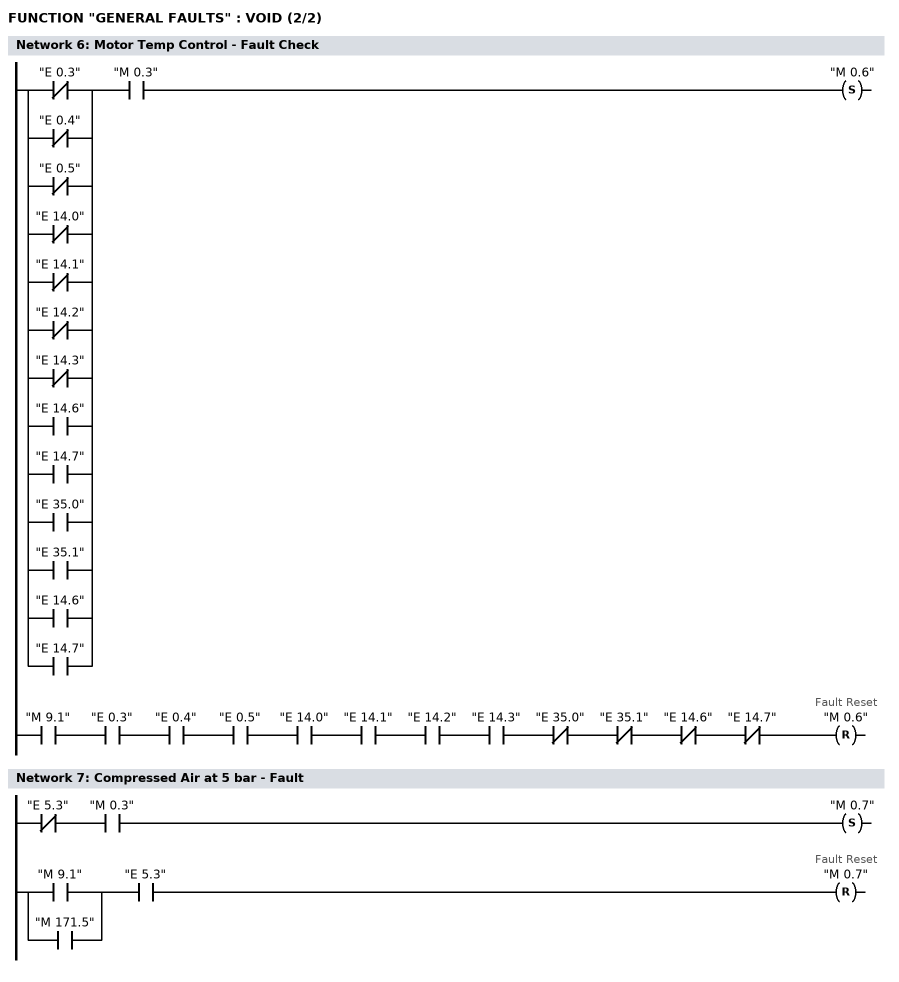

      A(    ;
      ON    "E 0.3";
      ON    "E 0.4";
      ON    "E 0.5";
      ON    "E 14.0";
      ON    "E 14.1";
      ON    "E 14.2";
      ON    "E 14.3";
      O     "E 14.6";
      O     "E 14.7";
      O     "E 35.0";
      O     "E 35.1";
      O     "E 14.6";
      O     "E 14.7";
      )     ;
      A     "M 0.3";
      S     "M 0.6";
//;
      A     "M 9.1";
      A     "E 0.3";
      A     "E 0.4";
      A     "E 0.5";
      A     "E 14.0";
      A     "E 14.1";
      A     "E 14.2";
      A     "E 14.3";
      AN    "E 35.0";
      AN    "E 35.1";
      AN    "E 14.6";
      AN    "E 14.7";
      R     "M 0.6"; // Fault Reset
NETWORK
TITLE =Compressed Air at 5 bar - Fault

      AN    "E 5.3";
      A     "M 0.3";
      S     "M 0.7";
//;
      A(    ;
      O     "M 9.1";
      O     "M 171.5";
      )     ;
      A     "E 5.3";
      R     "M 0.7"; // Fault Reset
NETWORK
TITLE =Faults Register 1 - E-Stops & Safety Doors

      A(    ;
      L     "MB 1";
      L     0;
      <>I   ;
      )     ;
      =     #FAULT_REGISTER_1;
//;
      A     #FAULT_REGISTER_1;
      O     #CHECK_PULSE;
      O     "M 17.1";
      O     "M 9.1";
      JNB   FR01;
NETWORK
TITLE =E-Stop  Desk  X120
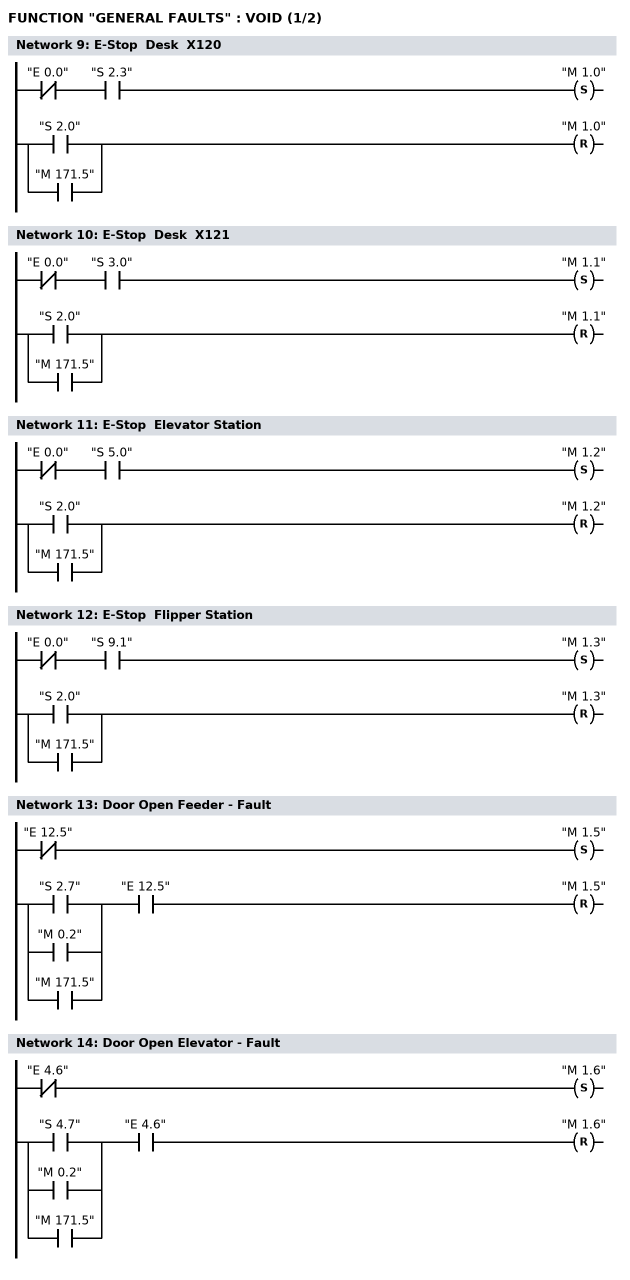

      AN    "E 0.0";
      A     "S 2.3";
      S     "M 1.0";
//;
      A(    ;
      O     "S 2.0";
      O     "M 171.5";
      )     ;
      R     "M 1.0";
NETWORK
TITLE =E-Stop  Desk  X121

      AN    "E 0.0";
      A     "S 3.0";
      S     "M 1.1";
//;
      A(    ;
      O     "S 2.0";
      O     "M 171.5";
      )     ;
      R     "M 1.1";
NETWORK
TITLE =E-Stop  Elevator Station

      AN    "E 0.0";
      A     "S 5.0";
      S     "M 1.2";
//;
      A(    ;
      O     "S 2.0";
      O     "M 171.5";
      )     ;
      R     "M 1.2";
NETWORK
TITLE =E-Stop  Flipper Station

      AN    "E 0.0";
      A     "S 9.1";
      S     "M 1.3";
//;
      A(    ;
      O     "S 2.0";
      O     "M 171.5";
      )     ;
      R     "M 1.3";
NETWORK
TITLE =Door Open Feeder - Fault

      AN    "E 12.5";
      S     "M 1.5";
//;
      A(    ;
      O     "S 2.7";
      O     "M 0.2";
      O     "M 171.5";
      )     ;
      A     "E 12.5";
      R     "M 1.5";
NETWORK
TITLE =Door Open Elevator - Fault

      AN    "E 4.6";
      S     "M 1.6";
//;
      A(    ;
      O     "S 4.7";
      O     "M 0.2";
      O     "M 171.5";
      )     ;
      A     "E 4.6";
      R     "M 1.6";
NETWORK
TITLE =Door Open Flipper - Fault
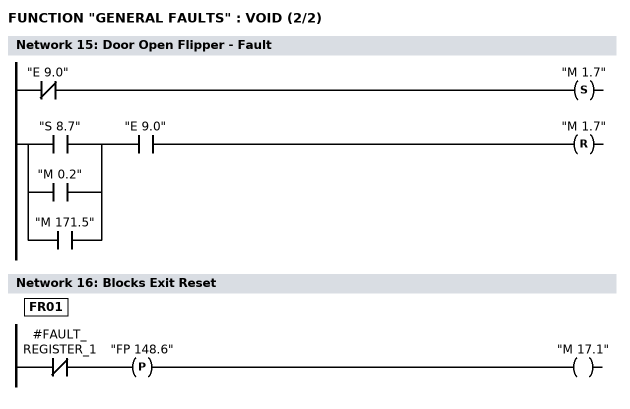

      AN    "E 9.0";
      S     "M 1.7";
//;
      A(    ;
      O     "S 8.7";
      O     "M 0.2";
      O     "M 171.5";
      )     ;
      A     "E 9.0";
      R     "M 1.7";
NETWORK
TITLE =Blocks Exit Reset

FR01: NOP   0;

      AN    #FAULT_REGISTER_1;
      FP    "FP 148.6";
      =     "M 17.1";
NETWORK
TITLE =Faults Register 2 - Conveyor 0 to Conveyor 3

      A(    ;
      L     "MB 2";
      L     0;
      <>I   ;
      )     ;
      =     #FAULT_REGISTER_2;
      =     "HMI_DB".SCREEN_CALL_1;
//;
      A     #FAULT_REGISTER_2;
      O     #CHECK_PULSE;
      O     "M 17.2";
      O     "M 9.1";
      JNB   FR02;
NETWORK
TITLE =K62.0 / 1 Conveyor 0 - Fault
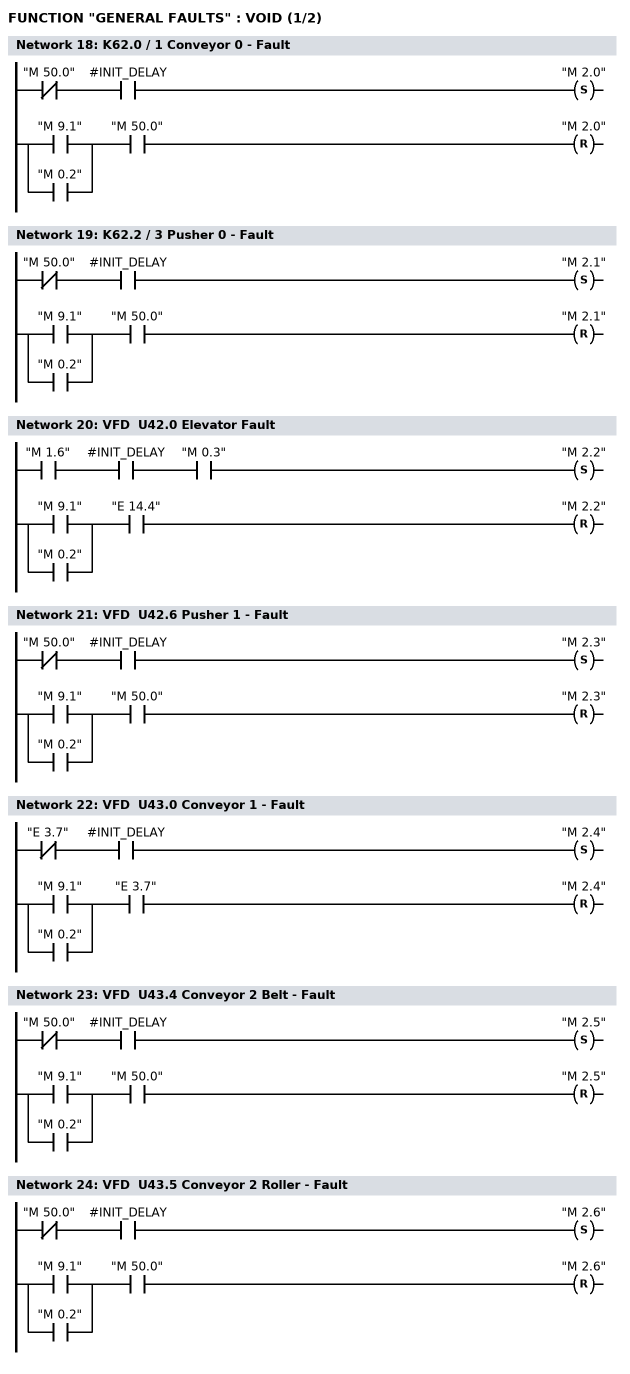

      AN    "M 50.0";
      A     #INIT_DELAY;
      S     "M 2.0";
//;
      A(    ;
      O     "M 9.1";
      O     "M 0.2";
      )     ;
      A     "M 50.0";
      R     "M 2.0";
NETWORK
TITLE =K62.2 / 3 Pusher 0 - Fault

      AN    "M 50.0";
      A     #INIT_DELAY;
      S     "M 2.1";
//;
      A(    ;
      O     "M 9.1";
      O     "M 0.2";
      )     ;
      A     "M 50.0";
      R     "M 2.1";
NETWORK
TITLE =VFD  U42.0 Elevator Fault

//   AN    #ELEVATOR_U42_0
      A     "M 1.6";
      A     #INIT_DELAY;
      A     "M 0.3";
      S     "M 2.2";
//;
      A(    ;
      O     "M 9.1";
      O     "M 0.2";
      )     ;
//      A     "E 3.6"
      A     "E 14.4";
      R     "M 2.2";
NETWORK
TITLE =VFD  U42.6 Pusher 1 - Fault

      AN    "M 50.0";
      A     #INIT_DELAY;
      S     "M 2.3";
//;
      A(    ;
      O     "M 9.1";
      O     "M 0.2";
      )     ;
      A     "M 50.0";
      R     "M 2.3";
NETWORK
TITLE =VFD  U43.0 Conveyor 1 - Fault

      AN    "E 3.7";
      A     #INIT_DELAY;
      S     "M 2.4";
//;
      A(    ;
      O     "M 9.1";
      O     "M 0.2";
      )     ;
      A     "E 3.7";
      R     "M 2.4";
NETWORK
TITLE =VFD  U43.4 Conveyor 2 Belt - Fault

      AN    "M 50.0";
      A     #INIT_DELAY;
      S     "M 2.5";
//;
      A(    ;
      O     "M 9.1";
      O     "M 0.2";
      )     ;
      A     "M 50.0";
      R     "M 2.5";
NETWORK
TITLE =VFD  U43.5 Conveyor 2 Roller - Fault

      AN    "M 50.0";
      A     #INIT_DELAY;
      S     "M 2.6";
//;
      A(    ;
      O     "M 9.1";
      O     "M 0.2";
      )     ;
      A     "M 50.0";
      R     "M 2.6";
NETWORK
TITLE =VFD  U44.0 Conveyor 3 Fault
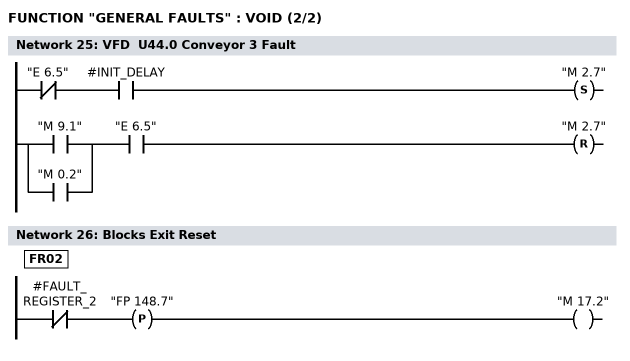

      AN    "E 6.5";
      A     #INIT_DELAY;
      S     "M 2.7";
//;
      A(    ;
      O     "M 9.1";
      O     "M 0.2";
      )     ;
      A     "E 6.5";
      R     "M 2.7";
NETWORK
TITLE =Blocks Exit Reset

FR02: NOP   0;

      AN    #FAULT_REGISTER_2;
      FP    "FP 148.7";
      =     "M 17.2";
NETWORK
TITLE =Faults Register 3 - Conveyor 4 to Conveyor 9

      A(    ;
      L     "MB 3";
      L     0;
      <>I   ;
      )     ;
      =     #FAULT_REGISTER_3;
      =     "HMI_DB".SCREEN_CALL_2;
//;
      A     #FAULT_REGISTER_3;
      O     #CHECK_PULSE;
      O     "M 17.3";
      O     "M 9.1";
      JNB   FR03;
NETWORK
TITLE =VFD  U44.3 Fault
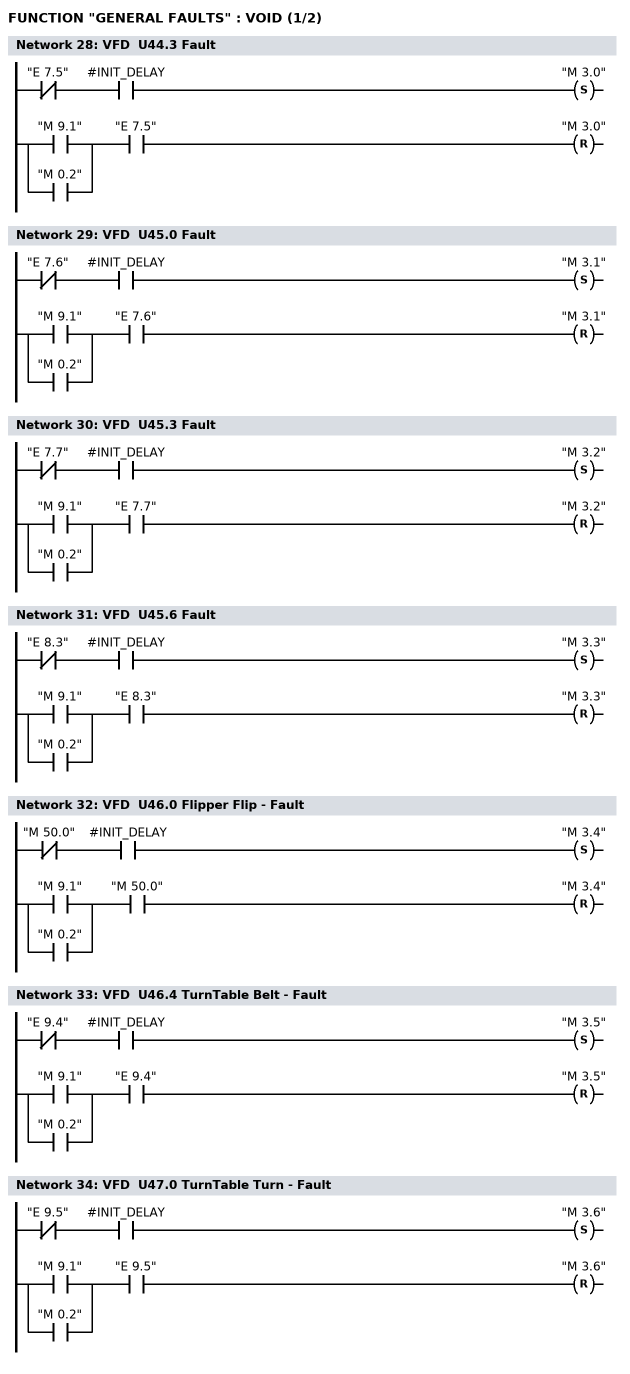

      AN    "E 7.5";
      A     #INIT_DELAY;
      S     "M 3.0";
//;
      A(    ;
      O     "M 9.1";
      O     "M 0.2";
      )     ;
      A     "E 7.5";
      R     "M 3.0";
NETWORK
TITLE =VFD  U45.0 Fault

      AN    "E 7.6";
      A     #INIT_DELAY;
      S     "M 3.1";
//;
      A(    ;
      O     "M 9.1";
      O     "M 0.2";
      )     ;
      A     "E 7.6";
      R     "M 3.1";
NETWORK
TITLE =VFD  U45.3 Fault

      AN    "E 7.7";
      A     #INIT_DELAY;
      S     "M 3.2";
//;
      A(    ;
      O     "M 9.1";
      O     "M 0.2";
      )     ;
      A     "E 7.7";
      R     "M 3.2";
NETWORK
TITLE =VFD  U45.6 Fault

      AN    "E 8.3";
      A     #INIT_DELAY;
      S     "M 3.3";
///;
      A(    ;
      O     "M 9.1";
      O     "M 0.2";
      )     ;
      A     "E 8.3";
      R     "M 3.3";
NETWORK
TITLE =VFD  U46.0 Flipper Flip - Fault

      AN    "M 50.0";
      A     #INIT_DELAY;
      S     "M 3.4";
//;
      A(    ;
      O     "M 9.1";
      O     "M 0.2";
      )     ;
      A     "M 50.0";
      R     "M 3.4";
NETWORK
TITLE =VFD  U46.4 TurnTable Belt - Fault

      AN    "E 9.4";
      A     #INIT_DELAY;
      S     "M 3.5";
//;
      A(    ;
      O     "M 9.1";
      O     "M 0.2";
      )     ;
      A     "E 9.4";
      R     "M 3.5";
NETWORK
TITLE =VFD  U47.0 TurnTable Turn - Fault

      AN    "E 9.5";
      A     #INIT_DELAY;
      S     "M 3.6";
//;
      A(    ;
      O     "M 9.1";
      O     "M 0.2";
      )     ;
      A     "E 9.5";
      R     "M 3.6";
NETWORK
TITLE =VFD  U47.5 Conveyor 9 - Fault
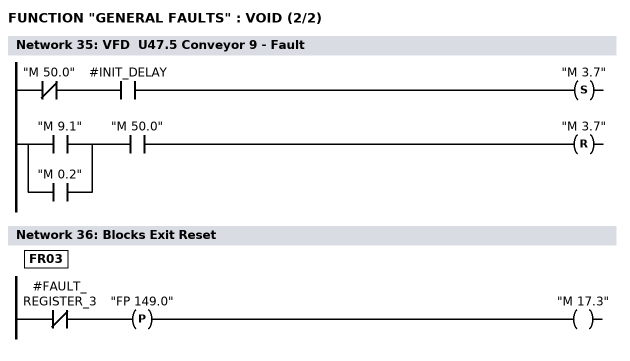

      AN    "M 50.0";
      A     #INIT_DELAY;
      S     "M 3.7";
//;
      A(    ;
      O     "M 9.1";
      O     "M 0.2";
      )     ;
      A     "M 50.0";
      R     "M 3.7";
NETWORK
TITLE =Blocks Exit Reset

FR03: NOP   0;

      AN    #FAULT_REGISTER_3;
      FP    "FP 149.0";
      =     "M 17.3";
NETWORK
TITLE =Faults Register 4 - Pusher 2 to Conveyor 23

      A(    ;
      L     "MB 4";
      L     0;
      <>I   ;
      )     ;
      =     #FAULT_REGISTER_4;
      =     "HMI_DB".SCREEN_CALL_2;
//;
      A     #FAULT_REGISTER_4;
      O     #CHECK_PULSE;
      O     "M 17.4";
      O     "M 9.1";
      JNB   FR04;
NETWORK
TITLE =VFD  U47.6 Pusher 2 - Fault
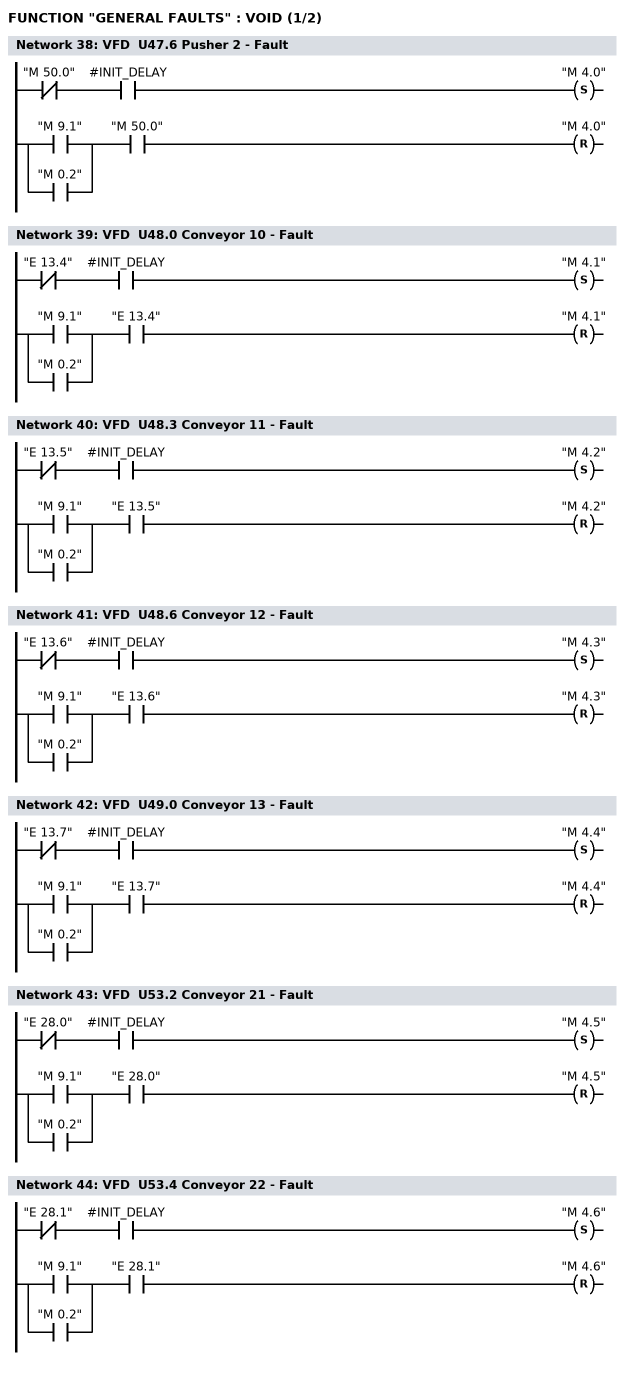

      AN    "M 50.0";
      A     #INIT_DELAY;
      S     "M 4.0";
//;
      A(    ;
      O     "M 9.1";
      O     "M 0.2";
      )     ;
      A     "M 50.0";
      R     "M 4.0";
NETWORK
TITLE =VFD  U48.0 Conveyor 10 - Fault

      AN    "E 13.4";
      A     #INIT_DELAY;
      S     "M 4.1";
//;
      A(    ;
      O     "M 9.1";
      O     "M 0.2";
      )     ;
      A     "E 13.4";
      R     "M 4.1";
NETWORK
TITLE =VFD  U48.3 Conveyor 11 - Fault

      AN    "E 13.5";
      A     #INIT_DELAY;
      S     "M 4.2";
//;
      A(    ;
      O     "M 9.1";
      O     "M 0.2";
      )     ;
      A     "E 13.5";
      R     "M 4.2";
NETWORK
TITLE =VFD  U48.6 Conveyor 12 - Fault

      AN    "E 13.6";
      A     #INIT_DELAY;
      S     "M 4.3";
//;
      A(    ;
      O     "M 9.1";
      O     "M 0.2";
      )     ;
      A     "E 13.6";
      R     "M 4.3";
NETWORK
TITLE =VFD  U49.0 Conveyor 13 - Fault

      AN    "E 13.7";
      A     #INIT_DELAY;
      S     "M 4.4";
//;
      A(    ;
      O     "M 9.1";
      O     "M 0.2";
      )     ;
      A     "E 13.7";
      R     "M 4.4";
NETWORK
TITLE =VFD  U53.2 Conveyor 21 - Fault

      AN    "E 28.0";
      A     #INIT_DELAY;
      S     "M 4.5";
//;
      A(    ;
      O     "M 9.1";
      O     "M 0.2";
      )     ;
      A     "E 28.0";
      R     "M 4.5";
NETWORK
TITLE =VFD  U53.4 Conveyor 22 - Fault

      AN    "E 28.1";
      A     #INIT_DELAY;
      S     "M 4.6";
//;
      A(    ;
      O     "M 9.1";
      O     "M 0.2";
      )     ;
      A     "E 28.1";
      R     "M 4.6";
NETWORK
TITLE =VFD  U54.0 Conveyor 23 - Fault
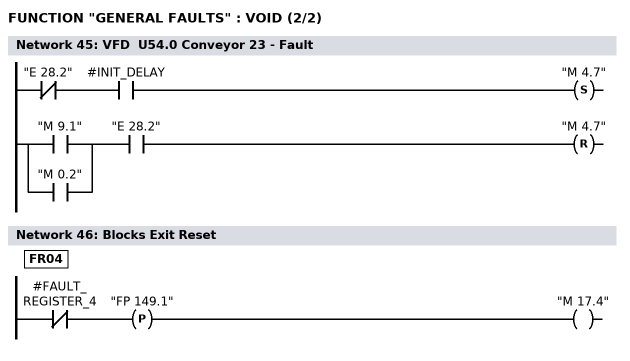

      AN    "E 28.2";
      A     #INIT_DELAY;
      S     "M 4.7";
//;
      A(    ;
      O     "M 9.1";
      O     "M 0.2";
      )     ;
      A     "E 28.2";
      R     "M 4.7";
NETWORK
TITLE =Blocks Exit Reset

FR04: NOP   0;

      AN    #FAULT_REGISTER_4;
      FP    "FP 149.1";
      =     "M 17.4";
NETWORK
TITLE =Faults Register 5 - Feeder

      A(    ;
      O     "M 7.0";
      O     "M 7.1";
      O     "M 7.2";
      )     ;
      =     #FAULT_REGISTER_5;
      =     "HMI_DB".SCREEN_CALL_3;
//;
      A     #FAULT_REGISTER_5;
      O     #CHECK_PULSE;
      O     "M 17.5";
      O     "M 9.1";
      JNB   FR05;
NETWORK
TITLE =VFD  U50.0 Feeder Lift - Fault
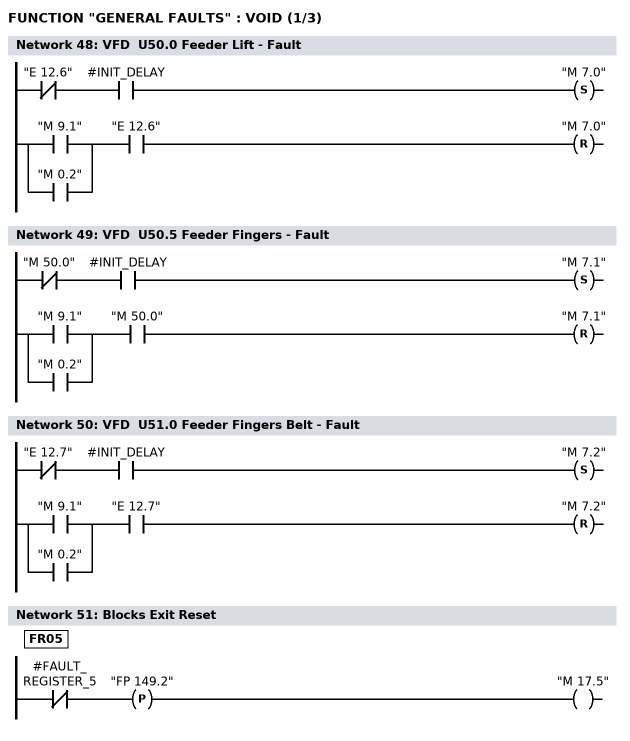

      AN    "E 12.6";
      A     #INIT_DELAY;
      S     "M 7.0";
//;
      A(    ;
      O     "M 9.1";
      O     "M 0.2";
      )     ;
      A     "E 12.6";
      R     "M 7.0";
NETWORK
TITLE =VFD  U50.5 Feeder Fingers - Fault

      AN    "M 50.0";
      A     #INIT_DELAY;
      S     "M 7.1";
//;
      A(    ;
      O     "M 9.1";
      O     "M 0.2";
      )     ;
      A     "M 50.0";
      R     "M 7.1";
NETWORK
TITLE =VFD  U51.0 Feeder Fingers Belt - Fault

      AN    "E 12.7";
      A     #INIT_DELAY;
      S     "M 7.2";
//;
      A(    ;
      O     "M 9.1";
      O     "M 0.2";
      )     ;
      A     "E 12.7";
      R     "M 7.2";
NETWORK
TITLE =Blocks Exit Reset

FR05: NOP   0;

      AN    #FAULT_REGISTER_5;
      FP    "FP 149.2";
      =     "M 17.5";
NETWORK
TITLE =Fault Status Lamp X120
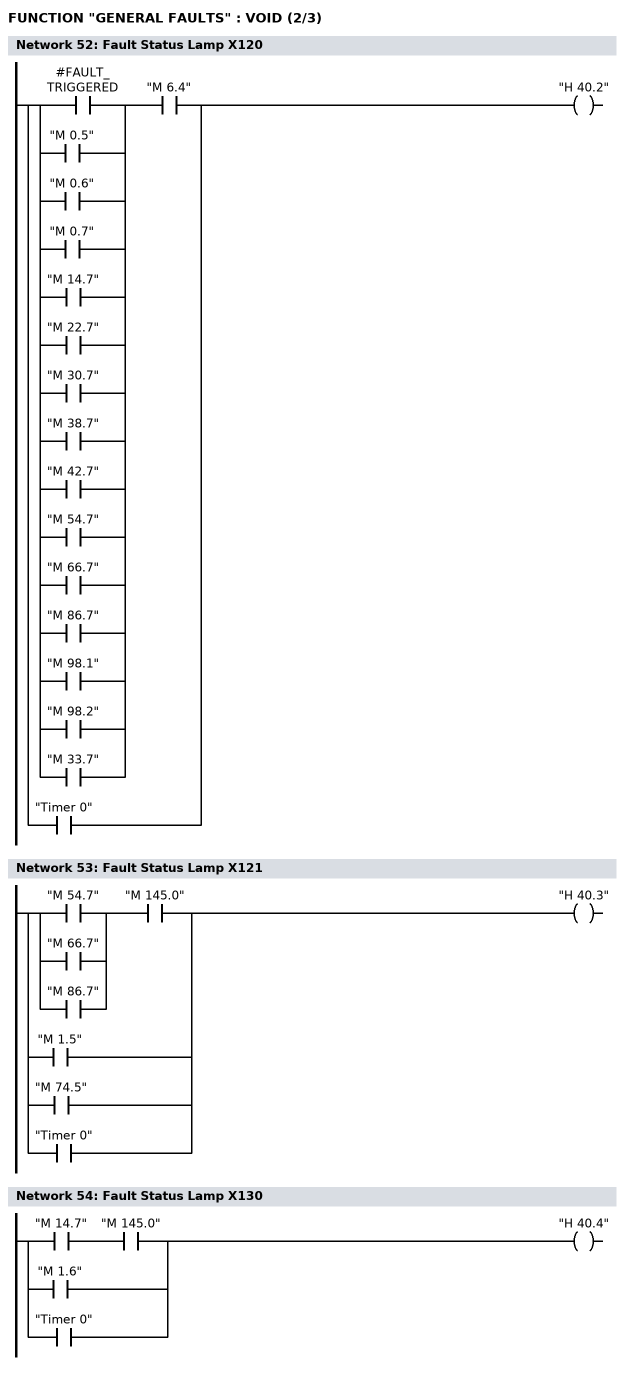

      A(    ;
      O     #FAULT_TRIGGERED;
      O     "M 0.5";
      O     "M 0.6";
      O     "M 0.7";
      O     "M 14.7";
      O     "M 22.7";
      O     "M 30.7";
      O     "M 38.7";
      O     "M 42.7";
      O     "M 54.7";
      O     "M 66.7";
      O     "M 86.7";
      O     "M 98.1";
      O     "M 98.2";
      O     "M 33.7";
      )     ;
      A     "M 6.4";
      O     "Timer 0";
      =     "H 40.2";
NETWORK
TITLE =Fault Status Lamp X121

      A(    ;
      O     "M 54.7";
      O     "M 66.7";
      O     "M 86.7";
      )     ;
      A     "M 145.0";
      O     "M 1.5";
      O     "M 74.5";
      O     "Timer 0";
      =     "H 40.3";
NETWORK
TITLE =Fault Status Lamp X130

      A     "M 14.7";
      A     "M 145.0";
      O     "M 1.6";
      O     "Timer 0";
      =     "H 40.4";
NETWORK
TITLE =Fault Status Lamp X134
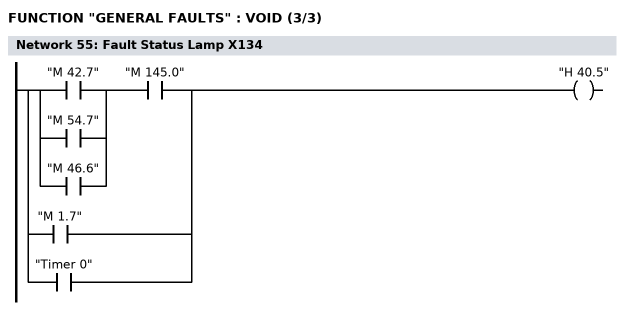

      A(    ;
      O     "M 42.7";
      O     "M 54.7";
      O     "M 46.6";
      )     ;
      A     "M 145.0";
      O     "M 1.7";
      O     "Timer 0";
      =     "H 40.5";
NETWORK
TITLE =Elevator OverTemp

      A     "M 0.6";
      AN    "E 0.3";
      L     W#16#1;
      T     "MB 181";
      BEC   ;
NETWORK
TITLE =Turntable OverTemp

      A     "M 0.6";
      AN    "E 0.4";
      L     W#16#2;
      T     "MB 181";
      BEC   ;
NETWORK
TITLE =Loader OverTemp

      A     "M 0.6";
      AN    "E 0.5";
      L     W#16#3;
      T     "MB 181";
      BEC   ;
NETWORK
TITLE =Conveyor 4 Collator OverTemp

      A     "M 0.6";
      AN    "E 14.0";
      L     W#16#4;
      T     "MB 181";
      BEC   ;
NETWORK
TITLE =Conveyor 6 Delivery OverTemp

      A     "M 0.6";
      AN    "E 14.1";
      L     W#16#5;
      T     "MB 181";
      BEC   ;
NETWORK
TITLE =Pivot Conveyor 10 OverTemp

      A(    ;
      ON    "E 14.2";
      ON    "E 14.3";
      )     ;
      A     "M 0.6";
      O     ;
      A(    ;
      O     "E 14.6";
      O     "E 14.7";
      )     ;
      A     "M 0.6";
      L     W#16#6;
      T     "MB 181";
      BEC   ;
NETWORK
TITLE =OverTemp

      A     "M 0.6";
      A     "E 35.0";
      L     W#16#8;
      T     "MB 181";
      BEC   ;
NETWORK
TITLE =OverTemp

      A     "M 0.6";
      A     "E 35.1";
      L     W#16#9;
      T     "MB 181";
      BEC   ;
NETWORK
TITLE =OverTemp

      A     "M 0.6";
      A     "E 14.6";
      L     W#16#B;
      T     "MB 181";
      BEC   ;
NETWORK
TITLE =OverTemp

      A     "M 0.6";
      A     "E 14.7";
      L     W#16#C;
      T     "MB 181";
      BEC   ;
NETWORK
TITLE =

      A     #FAULT_TRIGGERED;
      A     "M 3.0";
      L     W#16#0;
      T     MB   183;
      BEC   ;
NETWORK
TITLE =

      A     #FAULT_TRIGGERED;
      A     "M 3.1";
      L     W#16#1;
      T     MB   183;
      BEC   ;
NETWORK
TITLE =

      A     #FAULT_TRIGGERED;
      A     "M 3.2";
      L     W#16#2;
      T     MB   183;
      BEC   ;
NETWORK
TITLE =

      A     #FAULT_TRIGGERED;
      A     "M 3.3";
      L     W#16#3;
      T     MB   183;
      BEC   ;
NETWORK
TITLE =

      A     #FAULT_TRIGGERED;
      A     "M 3.4";
      L     W#16#4;
      T     MB   183;
      BEC   ;
NETWORK
TITLE =

      A     #FAULT_TRIGGERED;
      A     "M 3.5";
      L     W#16#5;
      T     MB   183;
      BEC   ;
NETWORK
TITLE =

      A     #FAULT_TRIGGERED;
      A     "M 3.6";
      L     W#16#6;
      T     MB   183;
      BEC   ;
NETWORK
TITLE =

      A     #FAULT_TRIGGERED;
      A     "M 3.7";
      L     W#16#7;
      T     MB   183;
      BEC   ;
NETWORK
TITLE =

      A     #FAULT_TRIGGERED;
      A     "M 4.0";
      L     W#16#8;
      T     MB   182;
      BEC   ;
NETWORK
TITLE =

      A     #FAULT_TRIGGERED;
      A     "M 4.1";
      L     W#16#9;
      T     MB   182;
      BEC   ;
NETWORK
TITLE =

      A     #FAULT_TRIGGERED;
      A     "M 4.2";
      L     W#16#10;
      T     MB   182;
      BEC   ;
NETWORK
TITLE =

      A     #FAULT_TRIGGERED;
      A     "M 4.3";
      L     W#16#11;
      T     MB   182;
      BEC   ;
NETWORK
TITLE =

      A     #FAULT_TRIGGERED;
      A     "M 4.4";
      L     W#16#12;
      T     MB   182;
      BEC   ;
NETWORK
TITLE =

      A     #FAULT_TRIGGERED;
      A     "M 4.5";
      L     W#16#13;
      T     MB   182;
      BEC   ;
NETWORK
TITLE =

      A     #FAULT_TRIGGERED;
      A     "M 4.6";
      L     W#16#14;
      T     MB   182;
      BEC   ;
NETWORK
TITLE =

      L     W#16#0;
      T     "MW 180";
      T     MW   182;
END_FUNCTION

FUNCTION "BLINKER" : VOID
TITLE =Blinker
VERSION : 0.0

BEGIN
NETWORK
TITLE =
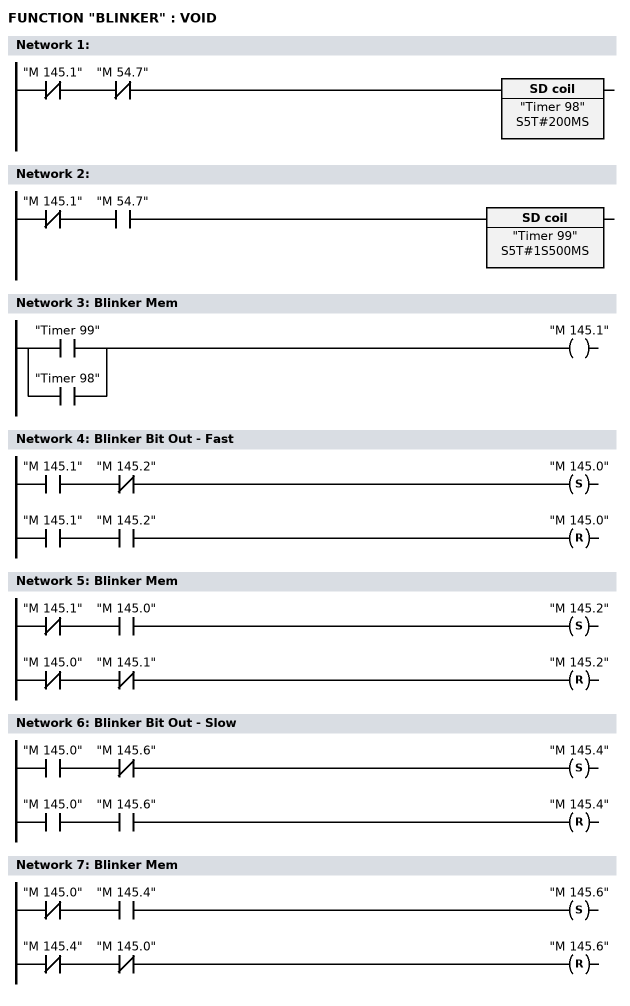

      AN    "M 145.1";
      AN    "M 54.7";
      L     S5T#200MS;
      SD    "Timer 98";
NETWORK
TITLE =

      AN    "M 145.1";
      A     "M 54.7";
      L     S5T#1S500MS;
      SD    "Timer 99";
NETWORK
TITLE =Blinker Mem

      O     "Timer 99";
      O     "Timer 98";
      =     "M 145.1";
NETWORK
TITLE =Blinker Bit Out - Fast

      A     "M 145.1";
      AN    "M 145.2";
      S     "M 145.0";
//;
      A     "M 145.1";
      A     "M 145.2";
      R     "M 145.0";
NETWORK
TITLE =Blinker Mem

      AN    "M 145.1";
      A     "M 145.0";
      S     "M 145.2";
//;
      AN    "M 145.0";
      AN    "M 145.1";
      R     "M 145.2";
NETWORK
TITLE =Blinker Bit Out - Slow

      A     "M 145.0";
      AN    "M 145.6";
      S     "M 145.4";
//;
      A     "M 145.0";
      A     "M 145.6";
      R     "M 145.4";
NETWORK
TITLE =Blinker Mem

      AN    "M 145.0";
      A     "M 145.4";
      S     "M 145.6";
//;
      AN    "M 145.4";
      AN    "M 145.0";
      R     "M 145.6";
END_FUNCTION

FUNCTION "LIGHT CURTAIN - SAFETY" : VOID
TITLE =Conveyors Catways - Access Safety
//Access to Conveyor 1-2-3 & 4 : Crossing Light Curtains Latches / Freezes these
//Conveyors !
//- To Resume Run, CatWay 1 (Conveyors 1-2-3) :  Push Top PB (Catway)
//and Push Lower PB (Main Floor) within 15sec .
//- To Resume Run, CatWay 2 (Conveyors 3-4) :  Push Top PB (Catway) .
//
//If Crossing CatWay 2 Light Curtain while No Conveyors are running, Run will
//resume automatic after 1 sec of free Light Curtain.
//
//Big Red Light will Blink to confirm the Conveyors are disabled / Safe .
VERSION : 0.1

BEGIN
NETWORK
TITLE =Safety Light Curtains -  Trigger 2 - Momentary SF = 1s
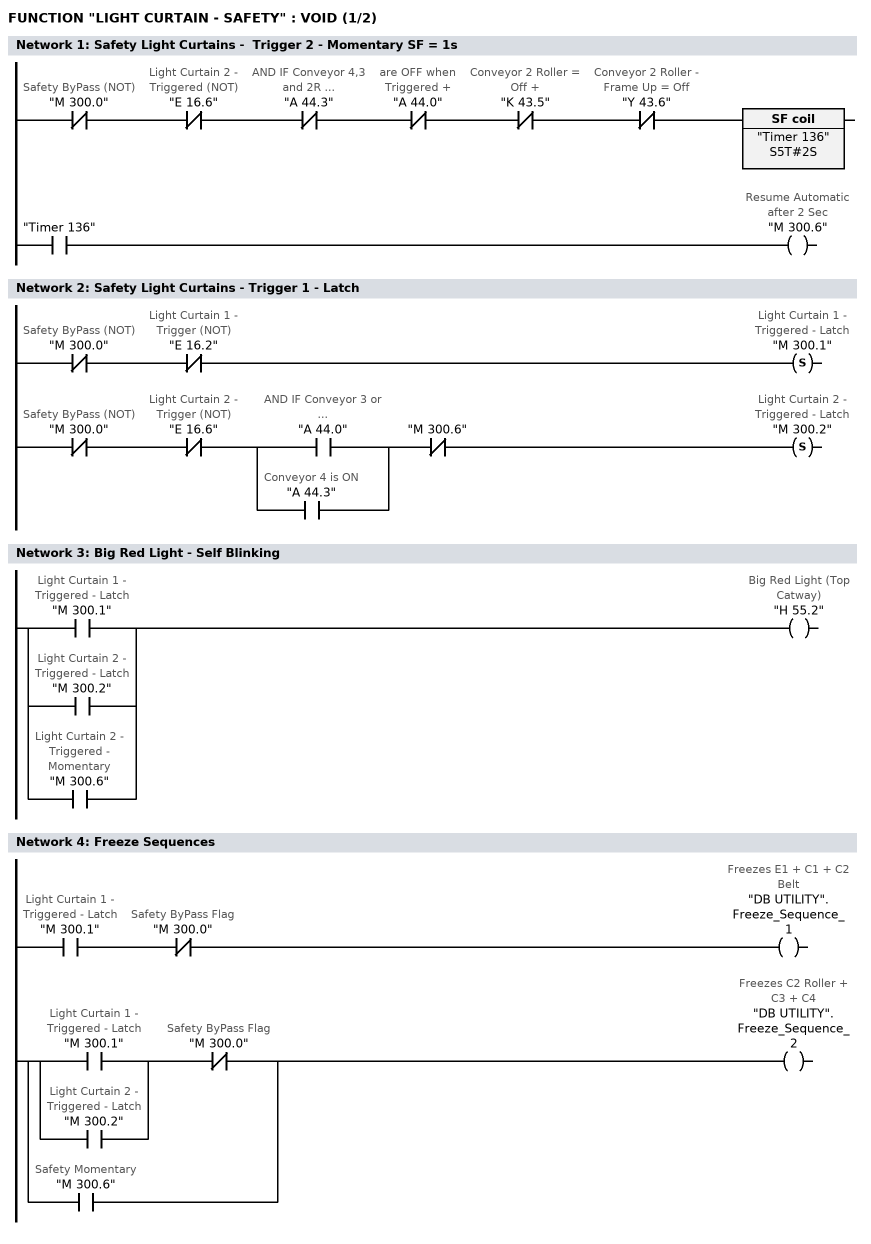

      AN    "M 300.0"; // Safety ByPass (NOT)
      AN    "E 16.6"; // Light Curtain 2 - Triggered (NOT)
      AN    "A 44.3"; // AND IF Conveyor 4,3 and 2R ...
      AN    "A 44.0"; // are OFF when Triggered +
      AN    "K 43.5"; // Conveyor 2 Roller = Off +
      AN    "Y 43.6"; // Conveyor 2 Roller - Frame Up = Off
      L     S5T#2S;
      SF    "Timer 136"; // Debouncer 2s
//;
      A     "Timer 136";
      =     "M 300.6"; // Resume Automatic after 2 Sec

NETWORK
TITLE =Safety Light Curtains - Trigger 1 - Latch

      AN    "M 300.0"; // Safety ByPass (NOT)
      AN    "E 16.2"; // Light Curtain 1 - Trigger (NOT)
      S     "M 300.1"; // Light Curtain 1 - Triggered - Latch
//;
      AN    "M 300.0"; // Safety ByPass (NOT)
      AN    "E 16.6"; // Light Curtain 2 - Trigger (NOT)
      A(    ;
      O     "A 44.0"; // AND IF Conveyor 3 or ...
      O     "A 44.3"; // Conveyor 4 is ON
      )     ;
      AN    "M 300.6";
      S     "M 300.2"; // Light Curtain 2 - Triggered - Latch
NETWORK
TITLE =Big Red Light - Self Blinking

      A(    ;
      O     "M 300.1"; // Light Curtain 1 - Triggered - Latch
      O     "M 300.2"; // Light Curtain 2 - Triggered - Latch
      O     "M 300.6"; // Light Curtain 2 - Triggered - Momentary
      )     ;
      =     "H 55.2"; // Big Red Light (Top Catway)
NETWORK
TITLE =Freeze Sequences

      A     "M 300.1"; // Light Curtain 1 - Triggered - Latch
      AN    "M 300.0"; // Safety ByPass Flag
      =     "DB UTILITY".Freeze_Sequence_1; //   Freezes E1 + C1 + C2 Belt
//;
      A     "M 300.1"; // Light Curtain 1 - Triggered - Latch
      O     "M 300.2"; // Light Curtain 2 - Triggered - Latch
      AN    "M 300.0"; // Safety ByPass Flag
      O     "M 300.6"; // Safety Momentary
      =     "DB UTILITY".Freeze_Sequence_2; //  Freezes C2 Roller + C3 + C4
NETWORK
TITLE =Safety ByPass - While blocking Curtain, Push Top Button for 5s
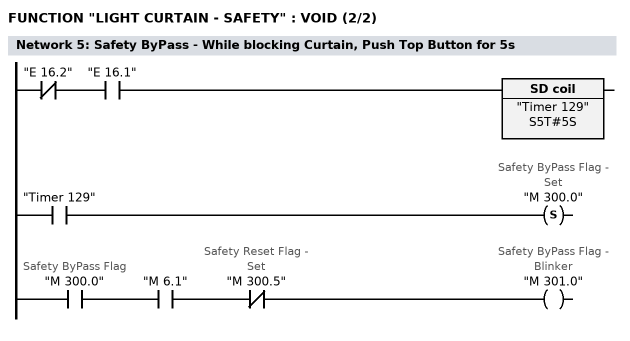

      AN    "E 16.2";
      A     "E 16.1";
      L     S5T#5S;
      SD    "Timer 129";
//;
      A     "Timer 129";
      S     "M 300.0"; // Safety ByPass Flag - Set
//;
      A     "M 300.0"; // Safety ByPass Flag
      A     "M 6.1";
      AN    "M 300.5"; // Safety Reset Flag - Set
      =     "M 301.0"; // Safety ByPass Flag - Blinker

NETWORK
TITLE =TEST REMOTE B+

      R     "A 58.4";

NETWORK
TITLE =PB Led - Control
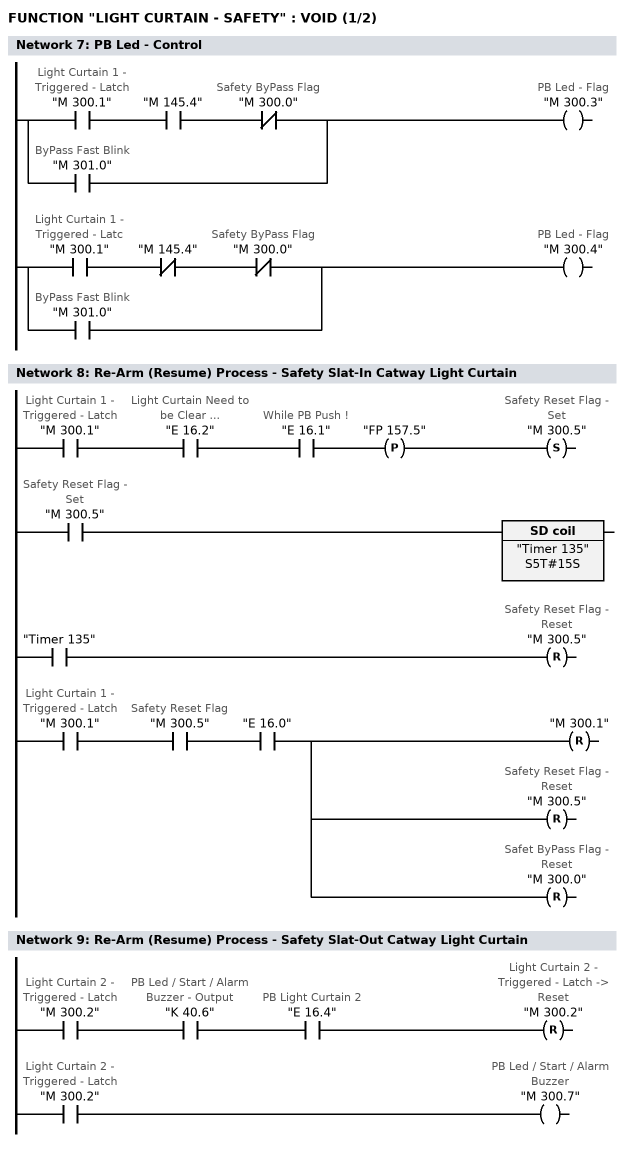

      A     "M 300.1"; // Light Curtain 1 - Triggered - Latch
      A     "M 145.4";
      AN    "M 300.0"; // Safety ByPass Flag
      O     "M 301.0"; // ByPass Fast Blink
      =     "M 300.3"; // PB Led - Flag
//;
      A     "M 300.1"; // Light Curtain 1 - Triggered - Latc
      AN    "M 145.4";
      AN    "M 300.0"; // Safety ByPass Flag
      O     "M 301.0"; // ByPass Fast Blink
      =     "M 300.4"; // PB Led - Flag
NETWORK
TITLE =Re-Arm (Resume) Process - Safety Slat-In Catway Light Curtain

      A     "M 300.1"; // Light Curtain 1 - Triggered - Latch
      A     "E 16.2"; // Light Curtain Need to be Clear ...
      A     "E 16.1"; // While PB Push !
      FP    "FP 157.5";
      S     "M 300.5"; // Safety Reset Flag - Set
//;
      A     "M 300.5"; // Safety Reset Flag - Set
      L     S5T#15S;
      SD    "Timer 135"; // Safety Reset Flag - TimeOut
//;
      A     "Timer 135";
      R     "M 300.5"; // Safety Reset Flag - Reset
//;
      A     "M 300.1"; // Light Curtain 1 - Triggered - Latch
      A     "M 300.5"; // Safety Reset Flag
      A     "E 16.0";
      R     "M 300.1";
      R     "M 300.5"; // Safety Reset Flag - Reset
      R     "M 300.0"; // Safet ByPass Flag - Reset
NETWORK
TITLE =Re-Arm (Resume) Process - Safety Slat-Out Catway Light Curtain

      A     "M 300.2"; // Light Curtain 2 - Triggered - Latch
      A     "K 40.6"; // PB Led / Start / Alarm Buzzer - Output
      A     "E 16.4"; // PB Light Curtain 2
      R     "M 300.2"; // Light Curtain 2 - Triggered - Latch -> Reset
//;
      A     "M 300.2"; // Light Curtain 2 - Triggered - Latch
      =     "M 300.7"; // PB Led / Start / Alarm Buzzer
NETWORK
TITLE =PB Led - Out
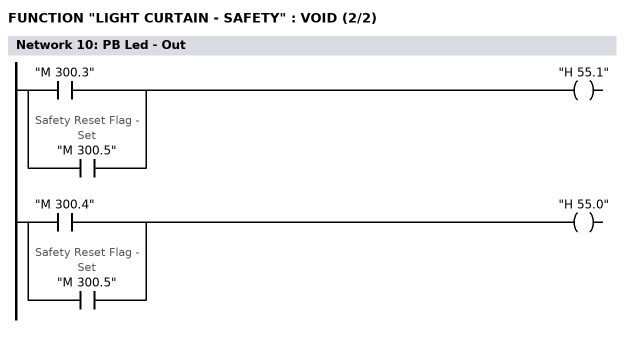

      A     "M 300.3";
      O     "M 300.5"; // Safety Reset Flag - Set
      =     "H 55.1";
//;
      A     "M 300.4";
      O     "M 300.5"; // Safety Reset Flag - Set
      =     "H 55.0";
END_FUNCTION

FUNCTION "NEW CLEARING" : VOID
TITLE =NEW FC911 (was FC1011) - Conveyors - Clearing Function
//New Order Sequence
//v0.1 2026-11-19: hold released at clearing start (FP M283.4); S3.2 lamp steady
//while held / blinking when ready; S3.2 held 3s releases the hold (T140).
NAME : CLEARING
VERSION : 0.1


VAR_TEMP
  EMPTY_11 : BOOL ;	//Empty Conveyor 11
  EMPTY_21 : BOOL ;	//Empty Conveyor 21
  EMPTY_12_22 : BOOL ;	//Empty Conveyor 12 & 22
  EMPTY_13_23 : BOOL ;	//Empty Conveyor 13 & 23
  C10_EMPTY_TEST : BOOL ;
  CLEARING_ABORT : BOOL ;
END_VAR
BEGIN
NETWORK
TITLE =HMI Clearing Call

      A     "M 140.3";
      A     "HMI_DB".CLEARING_SSW_MAIN;
      =     "M 5.2";
//;
      L     8;
      A     "M 10.0";
      =     "HMI_DB".CLEARING_SSW_STATUS;
      JC    CLEA;

      L     0;

CLEA: T     "HMI_DB".CLEARING_FUNCTION;

      A     "M 10.0";
      FN    "FN 155.7";
      R     "HMI_DB".CLEARING_SSW_MAIN;
      R     "M 54.2";
//;
      A     "M 5.2";
      FP    "FP 147.4";
      AN    "B 10.7"; // C11 - Empty
      AN    "B 11.0"; // C12 - Empty
      AN    "B 11.1"; // C13 - Empty
      AN    "B 11.2"; // C13 - Empty
      AN    "B 15.4"; // C21 - Empty
      AN    "B 15.5"; // C22 - Empty
      AN    "B 15.6"; // C23 - Empty
      AN    "B 15.7"; // C23 - Empty
      S     "M 54.2"; // Empty C11...C23
NETWORK
TITLE =New Order Seq - First New Order Packet to Pivot Conveyor 10
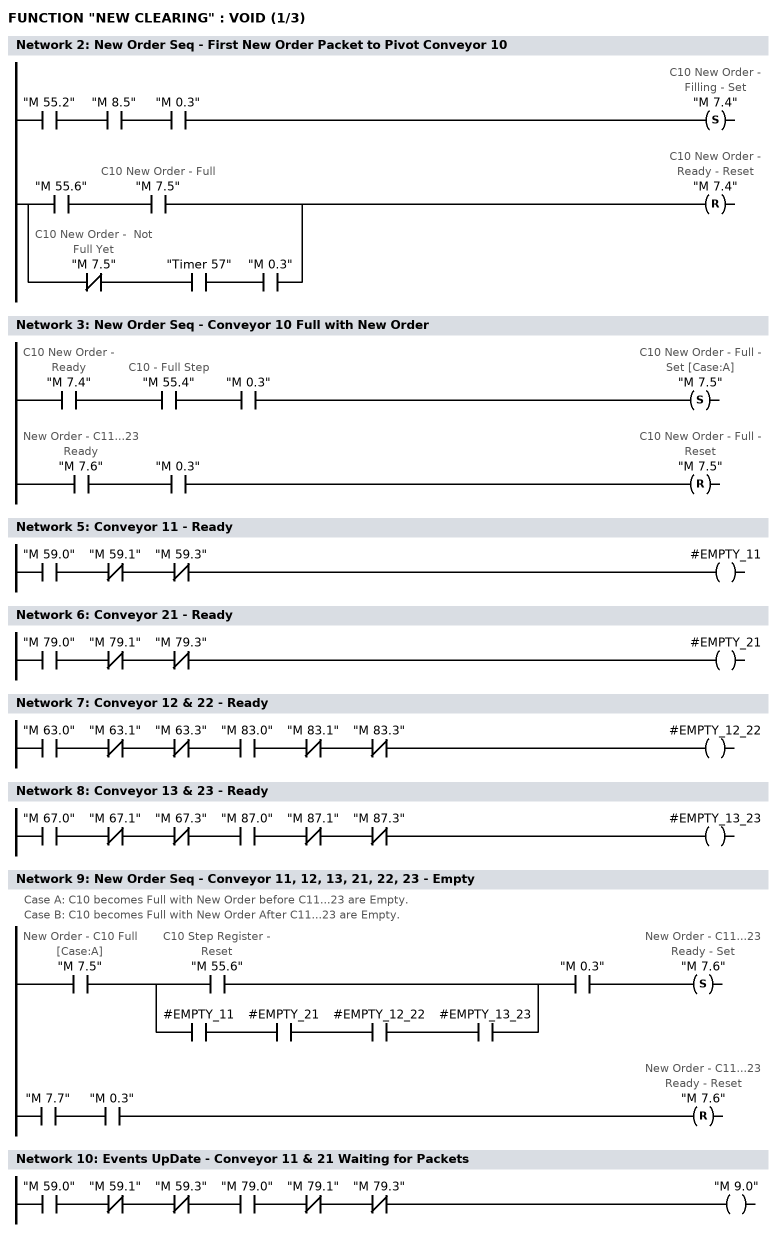

      A     "M 55.2";
      A     "M 8.5";
      A     "M 0.3";
      S     "M 7.4"; // C10 New Order - Filling - Set
//;
      A(    ;
      A     "M 55.6";
      A     "M 7.5"; // C10 New Order - Full
      O     ;
      AN    "M 7.5"; // C10 New Order -  Not Full Yet
      A     "Timer 57";
      A     "M 0.3";
      )     ;
      R     "M 7.4"; // C10 New Order - Ready - Reset
NETWORK
TITLE =New Order Seq - Conveyor 10 Full with New Order

      A     "M 7.4"; // C10 New Order - Ready
      A     "M 55.4"; // C10 - Full Step
      A     "M 0.3";
      S     "M 7.5"; // C10 New Order - Full - Set [Case:A]
//;
      A     "M 7.6"; // New Order - C11...23 Ready
      A     "M 0.3";
      R     "M 7.5"; // C10 New Order - Full - Reset
NETWORK
TITLE =New Order Seq
//New Order Seq - Waiting for the last Order Packets to Run out !


NETWORK
TITLE =Conveyor 11 - Ready

      A     "M 59.0";
      AN    "M 59.1";
      AN    "M 59.3";
      =     #EMPTY_11;
NETWORK
TITLE =Conveyor 21 - Ready

      A     "M 79.0";
      AN    "M 79.1";
      AN    "M 79.3";
      =     #EMPTY_21;
NETWORK
TITLE =Conveyor 12 & 22 - Ready

      A     "M 63.0";
      AN    "M 63.1";
      AN    "M 63.3";
      A     "M 83.0";
      AN    "M 83.1";
      AN    "M 83.3";
      =     #EMPTY_12_22;
NETWORK
TITLE =Conveyor 13 & 23 - Ready

      A     "M 67.0";
      AN    "M 67.1";
      AN    "M 67.3";
      A     "M 87.0";
      AN    "M 87.1";
      AN    "M 87.3";
      =     #EMPTY_13_23;
NETWORK
TITLE =New Order Seq - Conveyor 11, 12, 13, 21, 22, 23 - Empty
//Case A: C10 becomes Full with New Order before C11...23 are Empty.
//Case B: C10 becomes Full with New Order After C11...23 are Empty.
      A     "M 7.5"; // New Order - C10 Full [Case:A]
      A(    ;
      A     "M 55.6"; // C10 Step Register - Reset
      O     ;
      A     #EMPTY_11;
      A     #EMPTY_21;
      A     #EMPTY_12_22;
      A     #EMPTY_13_23;
      )     ;
      A     "M 0.3";
      S     "M 7.6"; // New Order - C11...23 Ready - Set
//;
      A     "M 7.7";
      A     "M 0.3";
      R     "M 7.6"; // New Order - C11...23 Ready - Reset
NETWORK
TITLE =Events UpDate - Conveyor 11 & 21 Waiting for Packets

      A     "M 59.0";
      AN    "M 59.1";
      AN    "M 59.3";
      A     "M 79.0";
      AN    "M 79.1";
      AN    "M 79.3";
      =     "M 9.0";
NETWORK
TITLE =New Order Seq - Conveyors 11, 21 - Empty
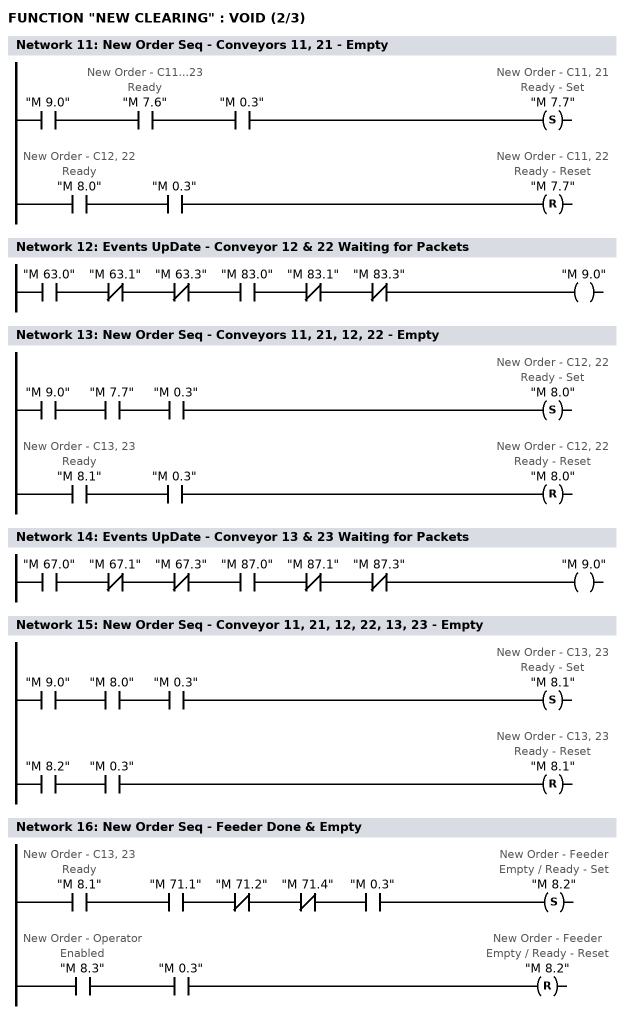

      A     "M 9.0";
      A     "M 7.6"; // New Order - C11...23 Ready
      A     "M 0.3";
      S     "M 7.7"; // New Order - C11, 21 Ready - Set
//;
      A     "M 8.0"; // New Order - C12, 22 Ready
      A     "M 0.3";
      R     "M 7.7"; // New Order - C11, 22 Ready - Reset
NETWORK
TITLE =Events UpDate - Conveyor 12 & 22 Waiting for Packets

      A     "M 63.0";
      AN    "M 63.1";
      AN    "M 63.3";
      A     "M 83.0";
      AN    "M 83.1";
      AN    "M 83.3";
      =     "M 9.0";
NETWORK
TITLE =New Order Seq - Conveyors 11, 21, 12, 22 - Empty

      A     "M 9.0";
      A     "M 7.7";
      A     "M 0.3";
      S     "M 8.0"; // New Order - C12, 22 Ready - Set
//;
      A     "M 8.1"; // New Order - C13, 23 Ready
      A     "M 0.3";
      R     "M 8.0"; // New Order - C12, 22 Ready - Reset
NETWORK
TITLE =Events UpDate - Conveyor 13 & 23 Waiting for Packets

      A     "M 67.0";
      AN    "M 67.1";
      AN    "M 67.3";
      A     "M 87.0";
      AN    "M 87.1";
      AN    "M 87.3";
      =     "M 9.0";
NETWORK
TITLE =New Order Seq - Conveyor 11, 21, 12, 22, 13, 23 - Empty

      A     "M 9.0";
      A     "M 8.0";
      A     "M 0.3";
      S     "M 8.1"; // New Order - C13, 23 Ready - Set
//;
      A     "M 8.2";
      A     "M 0.3";
      R     "M 8.1"; // New Order - C13, 23 Ready - Reset
NETWORK
TITLE =New Order Seq - Feeder Done & Empty

      A     "M 8.1"; // New Order - C13, 23 Ready
      A     "M 71.1";
      AN    "M 71.2";
      AN    "M 71.4";
      A     "M 0.3";
      S     "M 8.2"; // New Order - Feeder Empty / Ready - Set
//;
      A     "M 8.3"; // New Order - Operator Enabled
      A     "M 0.3";
      R     "M 8.2"; // New Order - Feeder Empty / Ready - Reset
NETWORK
TITLE =Conveyor 10 Clearing Enable after New Order
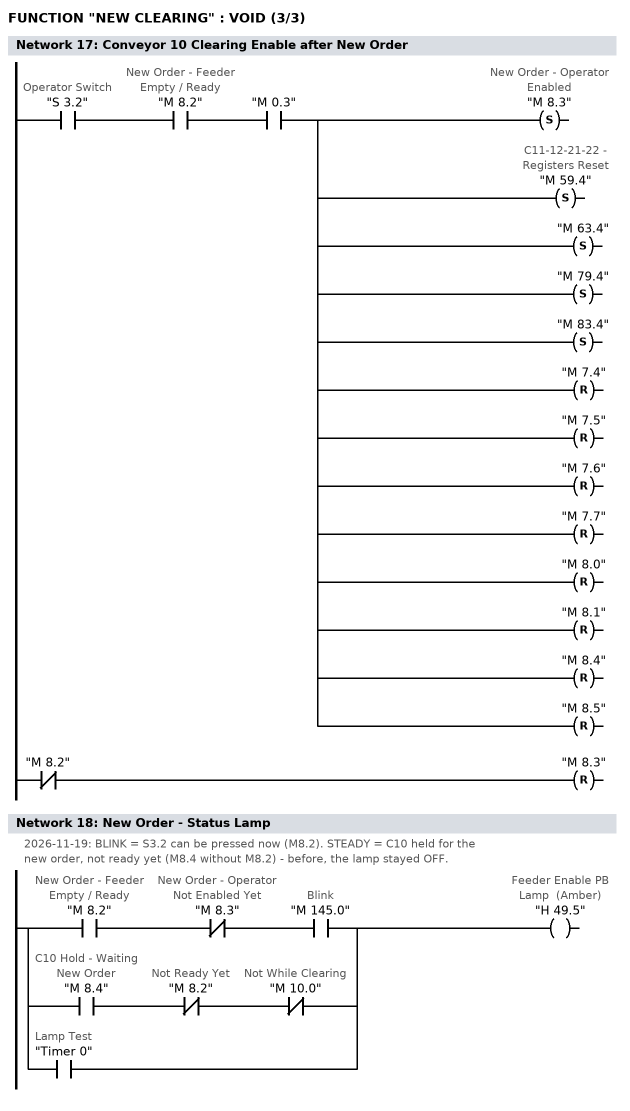

      A     "S 3.2"; // Operator Switch
      A     "M 8.2"; // New Order - Feeder Empty / Ready
      A     "M 0.3";
      S     "M 8.3"; // New Order - Operator Enabled
      S     "M 59.4"; // C11-12-21-22 - Registers Reset
      S     "M 63.4";
      S     "M 79.4";
      S     "M 83.4";
//;
      R     "M 7.4";
      R     "M 7.5";
      R     "M 7.6";
      R     "M 7.7";
      R     "M 8.0";
      R     "M 8.1";
      R     "M 8.4";
      R     "M 8.5";
//;
      ON    "M 8.2";
      R     "M 8.3";
NETWORK
TITLE =New Order - Status Lamp
//2026-11-19: BLINK = S3.2 can be pressed now (M8.2). STEADY = C10 held for the
//new order, not ready yet (M8.4 without M8.2) - before, the lamp stayed OFF.
      A(    ;
      A     "M 8.2"; // New Order - Feeder Empty / Ready
      AN    "M 8.3"; // New Order - Operator Not Enabled Yet
      A     "M 145.0"; // Blink
      )     ;
      O(    ;
      A     "M 8.4"; // C10 Hold - Waiting New Order
      AN    "M 8.2"; // Not Ready Yet
      AN    "M 10.0"; // Not While Clearing
      )     ;
      O     "Timer 0"; // Lamp Test
      =     "H 49.5"; // Feeder Enable PB Lamp  (Amber)
NETWORK
TITLE =S3.2 Held 3s - Release the Hold (Sequence Not Complete)
//2026-11-19: Before, S3.2 only worked with M8.2 (whole new-order chain done).
//If the chain got stuck, the TS waited with no way out but SIGNAL/F4.
//S3.2 held 3s releases the hold only (C11...C22 steps NOT reset: they may
//still carry the previous order).
      A     "S 3.2"; // Operator PB
      A     "M 8.4"; // C10 Hold Active
      AN    "M 10.0"; // Not While Clearing
      L     S5T#3S;
      SD    T    140; // Hold 3s (Free Timer)
//;
      A     T    140;
      A     "M 0.3";
      JCN   S321;

      R     "M 7.4";
      R     "M 7.5";
      R     "M 7.6";
      R     "M 7.7";
      R     "M 8.0";
      R     "M 8.1";
      R     "M 8.2";
      R     "M 8.3";
      R     "M 8.4"; // C10 Hold - Released
      R     "M 8.5"; // Clearing Done - Reset

S321: NOP   0;
NETWORK
TITLE =Conveyors Clearing Blink
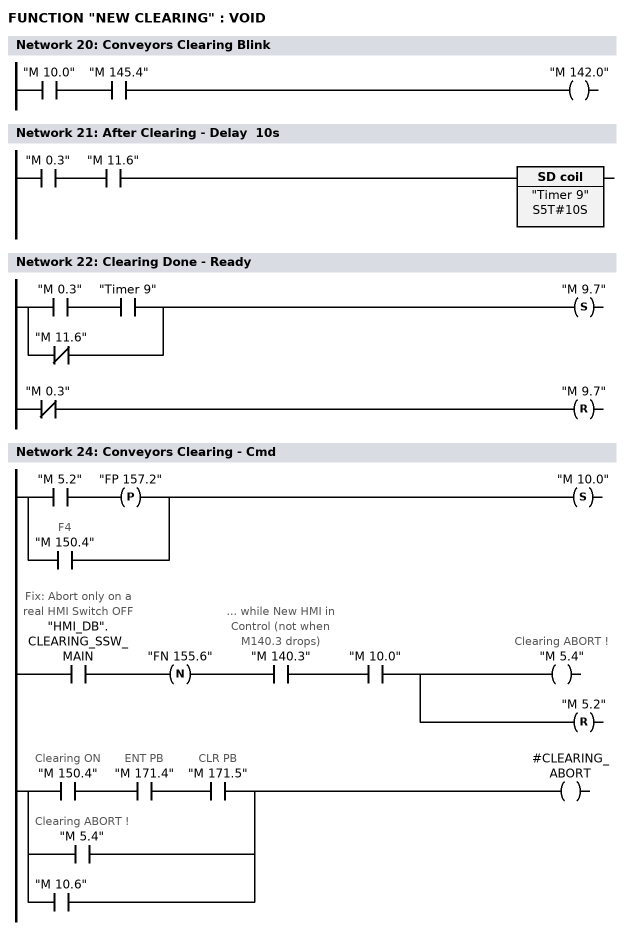

      A     "M 10.0";
      A     "M 145.4";
      =     "M 142.0";
NETWORK
TITLE =After Clearing - Delay  10s

      A     "M 0.3";
      A     "M 11.6";
      L     S5T#10S;
      SD    "Timer 9";
NETWORK
TITLE =Clearing Done - Ready

      A     "M 0.3";
      A     "Timer 9";
      ON    "M 11.6";
      S     "M 9.7";
//;
      ON    "M 0.3";
      R     "M 9.7";
NETWORK
TITLE =Clearing Command
//Clearing Command


NETWORK
TITLE =Conveyors Clearing - Cmd

      A(    ;
      A     "M 5.2";
      FP    "FP 157.2";
      O     ;
      A     "M 150.4"; // F4
      )     ;
      S     "M 10.0";
//;
      A     "HMI_DB".CLEARING_SSW_MAIN; // Fix: Abort only on a real HMI Switch OFF
      FN    "FN 155.6";
      A     "M 140.3"; // ... while New HMI in Control (not when M140.3 drops)
      A     "M 10.0";
      =     "M 5.4"; // Clearing ABORT !
      R     "M 5.2";
//;
      A(    ;
      A     "M 150.4"; // Clearing ON
      A     "M 171.4"; // ENT PB
      A     "M 171.5"; // CLR PB
      O     "M 5.4"; // Clearing ABORT !
      O     "M 10.6";
      )     ;
      =     #CLEARING_ABORT;
NETWORK
TITLE =Clearing Start - Release a Hold Left from the Previous Clearing
//Fix 2026-11-19: F4 pressed while C10 still held a new order (M8.4, S3.2 not
//pressed yet) -> C10 could not transfer, the clearing could never finish.
//F4 = clear everything: at every clearing start the hold and the new-order
//sequence are reset. They are set again when this clearing is done.
      A     "M 10.0"; // Clearing CMD
      FP    "FP 144.3"; // Edge Memory (Free)
      JCN   CST1;

      R     "M 7.4";
      R     "M 7.5";
      R     "M 7.6";
      R     "M 7.7";
      R     "M 8.0";
      R     "M 8.1";
      R     "M 8.2";
      R     "M 8.3";
      R     "M 8.4"; // C10 Hold - Released
      R     "M 8.5"; // Clearing Done - Reset

CST1: NOP   0;
NETWORK
TITLE =Conveyors Clearing Conveyors 1,2,3,4 - TimeOut 30S
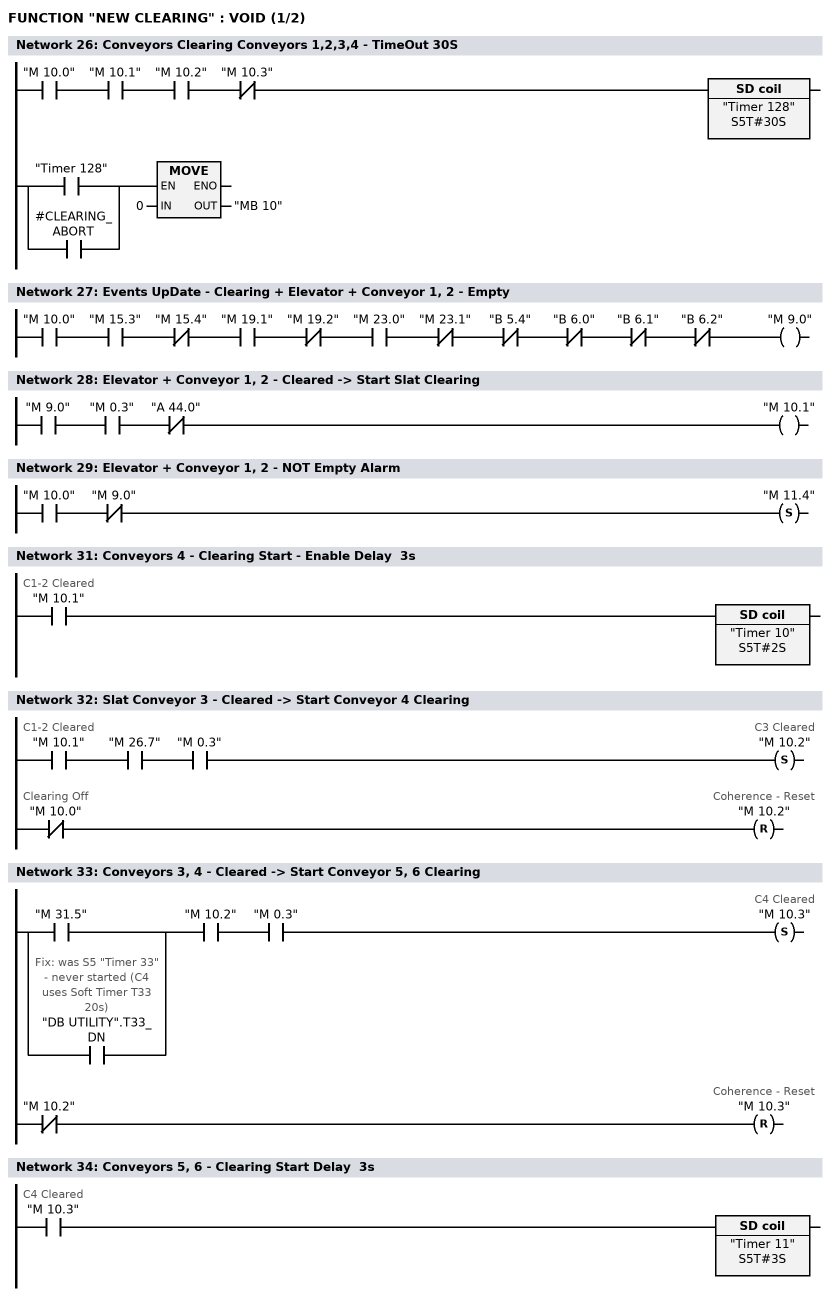

      A     "M 10.0";
      A     "M 10.1";
      A     "M 10.2";
      AN    "M 10.3";
      L     S5T#30S;
      SD    "Timer 128";
//;
      A     "Timer 128";
      O     #CLEARING_ABORT;
      JNB   NCLR;

      L     0;
      T     "MB 10"; // Clearing OFF

NCLR: NOP   0;
NETWORK
TITLE =Events UpDate - Clearing + Elevator + Conveyor 1, 2 - Empty

      A     "M 10.0";
      A     "M 15.3";
      AN    "M 15.4";
      A     "M 19.1";
      AN    "M 19.2";
      A     "M 23.0";
      AN    "M 23.1";
      AN    "B 5.4";
      AN    "B 6.0";
      AN    "B 6.1";
      AN    "B 6.2";
      =     "M 9.0";
NETWORK
TITLE =Elevator + Conveyor 1, 2 - Cleared -> Start Slat Clearing

      A     "M 9.0";
      A     "M 0.3";
      AN    "A 44.0";
      =     "M 10.1";
NETWORK
TITLE =Elevator + Conveyor 1, 2 - NOT Empty Alarm

      A     "M 10.0";
      AN    "M 9.0";
      S     "M 11.4";
NETWORK
TITLE =Clearing Sequence
//Clearing Sequence from Slat 3 to Pivot 10 Conveyors


NETWORK
TITLE =Conveyors 4 - Clearing Start - Enable Delay  3s

      A     "M 10.1"; // C1-2 Cleared
      L     S5T#2S;
      SD    "Timer 10";
NETWORK
TITLE =Slat Conveyor 3 - Cleared -> Start Conveyor 4 Clearing

      A     "M 10.1"; // C1-2 Cleared
      A     "M 26.7";
      A     "M 0.3";
      S     "M 10.2"; // C3 Cleared
//;
      AN    "M 10.0"; // Clearing Off
      R     "M 10.2"; // Coherence - Reset
NETWORK
TITLE =Conveyors 3, 4 - Cleared -> Start Conveyor 5, 6 Clearing

      A(    ;
      O     "M 31.5";
      O     "DB UTILITY".T33_DN; // Fix: was S5 "Timer 33" - never started (C4 uses Soft Timer T33 20s)
      )     ;
      A     "M 10.2";
      A     "M 0.3";
      S     "M 10.3"; // C4 Cleared
//;
      AN    "M 10.2";
      R     "M 10.3"; // Coherence - Reset
NETWORK
TITLE =Conveyors 5, 6 - Clearing Start Delay  3s

      A     "M 10.3"; // C4 Cleared
      L     S5T#3S;
      SD    "Timer 11"; // C4 Cleared Delayed
NETWORK
TITLE =Events UpDate - Conveyors 5, 6 - Clearing
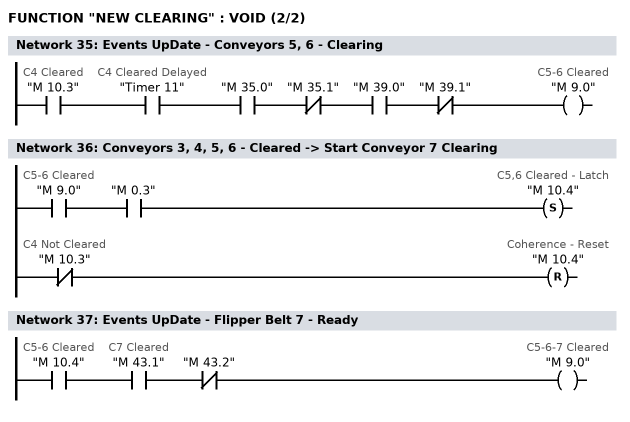

      A     "M 10.3"; // C4 Cleared
      A     "Timer 11"; // C4 Cleared Delayed
      A     "M 35.0";
      AN    "M 35.1";
      A     "M 39.0";
      AN    "M 39.1";
      =     "M 9.0"; // C5-6 Cleared
NETWORK
TITLE =Conveyors 3, 4, 5, 6 - Cleared -> Start Conveyor 7 Clearing

      A     "M 9.0"; // C5-6 Cleared
      A     "M 0.3";
      S     "M 10.4"; // C5,6 Cleared - Latch
//;
      AN    "M 10.3"; // C4 Not Cleared
      R     "M 10.4"; // Coherence - Reset
NETWORK
TITLE =Events UpDate - Flipper Belt 7 - Ready

      A     "M 10.4"; // C5-6 Cleared
      A     "M 43.1"; // C7 Cleared
      AN    "M 43.2";
      =     "M 9.0"; // C5-6-7 Cleared
NETWORK
TITLE =Conveyors 3, 4, 5, 6, 7, 8, 9 - Clearing - Cleared / Ready

      A     "M 9.0"; // C5-6-7 Cleared
      A     "M 47.2"; // C8 Cleared
      AN    "M 47.3";
      A     "M 51.1"; // C9 Cleared
      AN    "M 51.2";
      AN    "B 9.7"; // C9 - Pusher2 - Edge Cleared
      A     "M 0.3";
      L     S5T#3S;
      SD    "Timer 56"; // Delay 3s
//;
      A     "Timer 56";
      =     "M 10.5"; // C10 UpStream Cleared
      FP    "M 188.4";
      S     "M 58.2"; // C10 UpStream Cleared - Trigger Set
//;
      A     "M 10.5";
      L     S5T#1S;
      SE    "Timer 58"; // UpStream Cleared - Pulse 1s
NETWORK
TITLE =Clearing - C10 Proven Empty (Exit Sens Clear While Belt Runs Fas
//Fix: Clearing used to end with packets left on C10 (nothing checked C10 itself).
//C10 is proven empty when its Exit Sens B10.6 stays clear while the belt runs
//FAST (transfer) for the time a packet needs to cross the whole belt.
//TUNE: C10 belt length / 0.52 m/s (31 m/min) + margin.  10s = about 5 m.
//Any packet seen on C10 (B10.3 / B10.4 / B10.5 / B10.6) or a Pusher 2 push
//cancels the proof (a pushed packet can sit at the infeed without C10 starting).
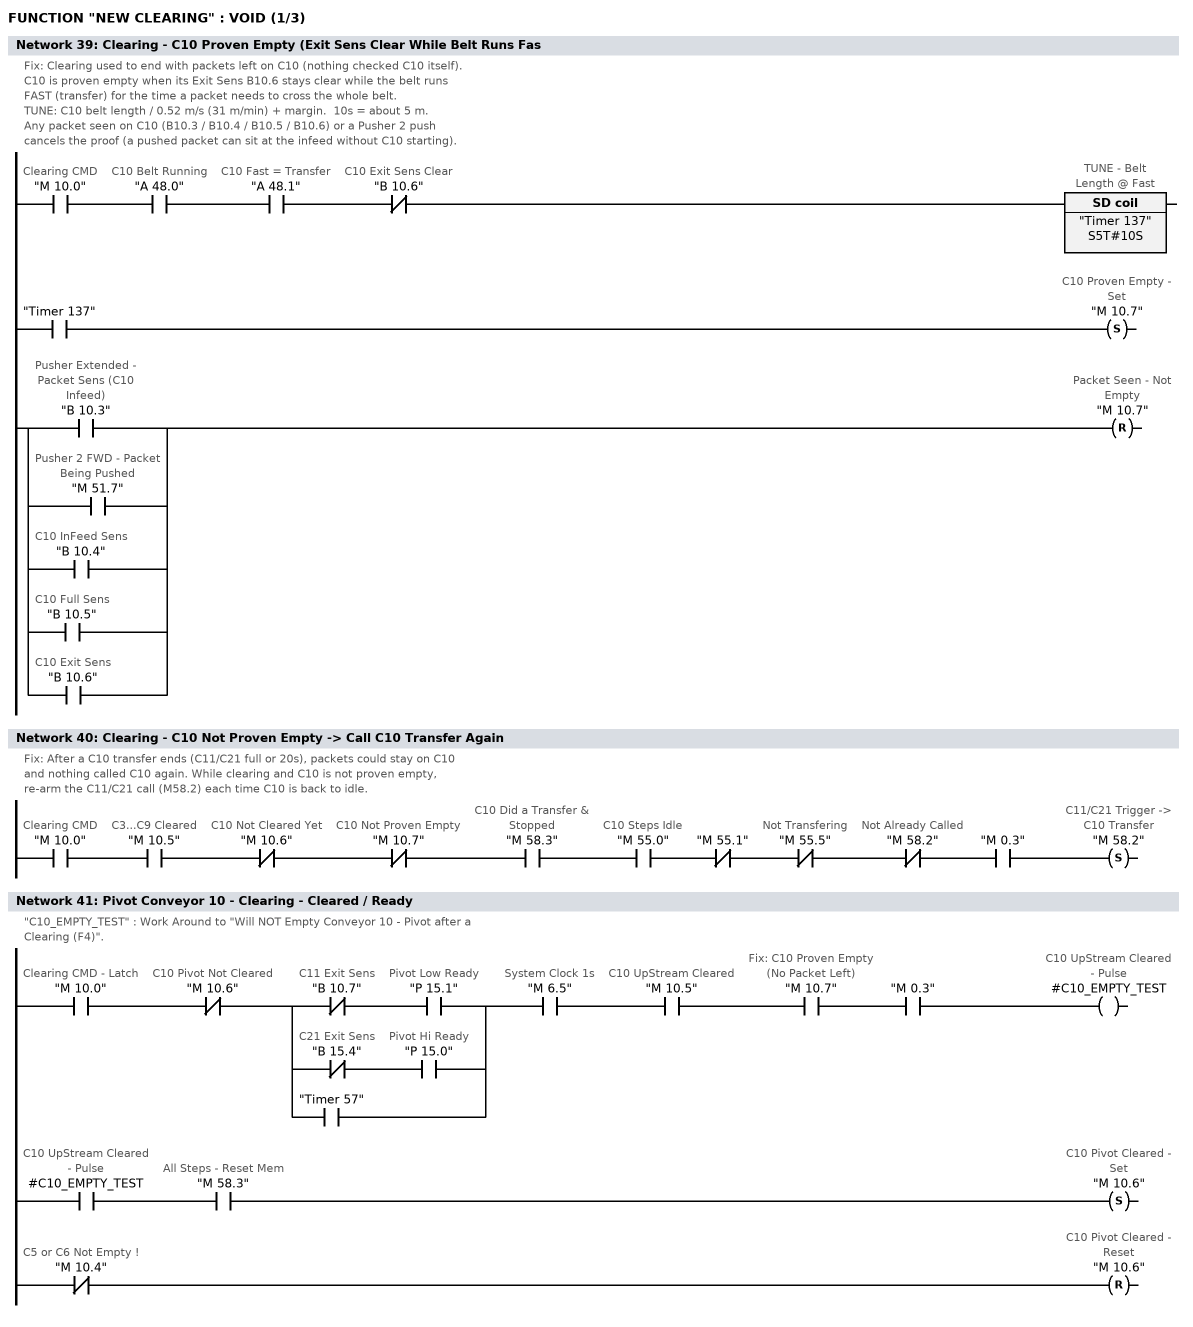
      A     "M 10.0"; // Clearing CMD
      A     "A 48.0"; // C10 Belt Running
      A     "A 48.1"; // C10 Fast = Transfer
      AN    "B 10.6"; // C10 Exit Sens Clear
      L     S5T#10S; // TUNE - Belt Length @ Fast
      SD    "Timer 137";
//;
      A     "Timer 137";
      S     "M 10.7"; // C10 Proven Empty - Set
//;
      A(    ;
      O     "B 10.3"; // Pusher Extended - Packet Sens (C10 Infeed)
      O     "M 51.7"; // Pusher 2 FWD - Packet Being Pushed
      O     "B 10.4"; // C10 InFeed Sens
      O     "B 10.5"; // C10 Full Sens
      O     "B 10.6"; // C10 Exit Sens
      )     ;
      R     "M 10.7"; // Packet Seen - Not Empty
NETWORK
TITLE =Clearing - C10 Not Proven Empty -> Call C10 Transfer Again
//Fix: After a C10 transfer ends (C11/C21 full or 20s), packets could stay on C10
//and nothing called C10 again. While clearing and C10 is not proven empty,
//re-arm the C11/C21 call (M58.2) each time C10 is back to idle.
      A     "M 10.0"; // Clearing CMD
      A     "M 10.5"; // C3...C9 Cleared
      AN    "M 10.6"; // C10 Not Cleared Yet
      AN    "M 10.7"; // C10 Not Proven Empty
      A     "M 58.3"; // C10 Did a Transfer & Stopped
      A     "M 55.0"; // C10 Steps Idle
      AN    "M 55.1";
      AN    "M 55.5"; // Not Transfering
      AN    "M 58.2"; // Not Already Called
      A     "M 0.3";
      S     "M 58.2"; // C11/C21 Trigger -> C10 Transfer
NETWORK
TITLE =Pivot Conveyor 10 - Clearing - Cleared / Ready
//"C10_EMPTY_TEST" : Work Around to "Will NOT Empty Conveyor 10 - Pivot after a
//Clearing (F4)".
      A     "M 10.0"; // Clearing CMD - Latch
      AN    "M 10.6"; // C10 Pivot Not Cleared
      A(    ;
      AN    "B 10.7"; // C11 Exit Sens
      A     "P 15.1"; // Pivot Low Ready
      O     ;
      AN    "B 15.4"; // C21 Exit Sens
      A     "P 15.0"; // Pivot Hi Ready
      O     "Timer 57";
      )     ;
      A     "M 6.5"; // System Clock 1s
      A     "M 10.5"; // C10 UpStream Cleared
      A     "M 10.7"; // Fix: C10 Proven Empty (No Packet Left)
      A     "M 0.3";
      =     #C10_EMPTY_TEST; // C10 UpStream Cleared - Pulse
//;
      A     #C10_EMPTY_TEST; // C10 UpStream Cleared - Pulse
      A     "M 58.3"; // All Steps - Reset Mem
      S     "M 10.6"; // C10 Pivot Cleared - Set
//;
      AN    "M 10.4"; // C5 or C6 Not Empty !
      R     "M 10.6"; // C10 Pivot Cleared - Reset
NETWORK
TITLE =C10 Clearing Trigger via C11 or C21
